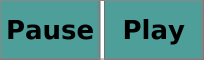
VISUALIZATION OperationButtons  // 204x60
VAR_IN_OUT
	stOperation	:ST_OperationButtons;
END_VAR
    Button (0,0 100x60), "Pause", tooltip "%s", colour toggle: stOperation.iActOperation=ePauseAll
        p4168582468: stOperation.sModeZone
        OnMouseClick: execute { stOperation.bSetPause:=TRUE; stOperation.iPauseHistory:=7; }
    Button (104,0 100x60), "Play", tooltip "%s", colour toggle: stOperation.iActOperation=ePlayAll
        p4168582468: stOperation.sModeZone
        OnMouseClick: execute { stOperation.bSetPlay:=TRUE; }
END_VISUALIZATION

(* stored: Version 1.1.0.1, ProductVersion 3.1.4024.13
   Visu OperationButtons: Id {fdcb95b3-d734-467c-9775-45181d98d290} *)
